Fanuc KAREL source: ka00132.KL

-- PROVISIONAL review KL for V1013-1; original PC SHA256 8da54f16c74d71c7e84ef2bb46fdd0d7e7532d247fc67e4dce6dcdc914fdbe91
-- Incomplete behavior may be omitted. Consult companion uncertainty JSON. Do not deploy.
PROGRAM KA00132
%NOLOCKGROUP
-- UNRESOLVED_DECL SRC type=002018
-- UNRESOLVED_DECL DST type=002017
BEGIN
  -- UNRESOLVED_PC offsets 5-19; opcodes 2E,22,9D,33,B2
  -- UNRESOLVED_PC offsets 24-42; opcodes 22,9D,33,B1,22,9D,33,B4
  -- UNRESOLVED_PC offsets 47-51; opcodes 7F
END KA00132
